Fanuc KAREL source: kt00450.KL

-- PROVISIONAL review KL for V770-1; original PC SHA256 91e1d367e2565b91e9e3e9ff64162ba0aed9e9b095dd2bb1934c9d6ef24b9b80
-- Incomplete behavior may be omitted. Consult companion uncertainty JSON. Do not deploy.
PROGRAM KT00450
%NOLOCKGROUP
VAR
  OUT : BOOLEAN
-- UNRESOLVED_DECL Y1 type=002018
-- UNRESOLVED_DECL H2 type=002017
BEGIN
  -- UNRESOLVED_PC offsets 5-19; opcodes 2E,22,9D,33,B2
  -- UNRESOLVED_PC offsets 24-38; opcodes 2E,22,9D,33,B4
  -- UNRESOLVED_PC offsets 43-68; opcodes 22,9D,33,B1,22,9D,33,B3,5C,23
  -- UNRESOLVED_PC offsets 73-77; opcodes 7F
END KT00450
